Fanuc KAREL source: ka00090.KL

PROGRAM KA00090
%STACKSIZE=65535
%PRIORITY=65535
%NOLOCKGROUP
VAR
SRC : JOINTPOS9
DST : XYZWPR
BEGIN
-- UNSAFE_SOURCE_IR line 7: DST = convert_jointpos9_to_xyzwpr(SRC)
END KA00090
